(* IEC 61131-3 sources: ZPLC/tools/hil/il_tests, 12 files *)

(* ---- arithmetic.il ---- *)
PROGRAM Arithmetic
VAR
  a AT %QW0 : INT;
  b AT %QW1 : INT;
  res_add AT %QW2 : INT;
  res_sub AT %QW3 : INT;
  res_mul AT %QW4 : INT;
  res_div AT %QW5 : INT;
  res_mod AT %QW6 : INT;
END_VAR

(* Explicit init for test stability *)
LD 10
ST a
LD 5
ST b

LD a
ADD b
ST res_add
LD a
SUB b
ST res_sub
LD a
MUL b
ST res_mul
LD a
DIV b
ST res_div
LD a
MOD b
ST res_mod
END_PROGRAM

(* ---- basic_il.il ---- *)
PROGRAM ILTest
VAR
    a AT %QW0 : INT := 10;
    b AT %QW1 : INT := 20;
    res AT %QW2 : INT;
    flag AT %QX6.0 : BOOL;
END_VAR

LD a
ADD b
ST res

LD res
GT 25
ST flag

END_PROGRAM

(* ---- blinky.il ---- *)
PROGRAM BlinkIL
VAR
  Blink : TON;
  Led AT %QX0.0 : BOOL;
END_VAR

(* The timer runs while the LED is off. When it is done the LED is on for one scan, which restarts the timer. *)
  LDN Led
  ST Blink.IN
  CAL Blink(PT := T#200ms)
  LD Blink.Q
  ST Led
END_PROGRAM

(* ---- comparison.il ---- *)
PROGRAM Comparison
VAR
  val AT %QW0 : INT;
  is_gt AT %QX2.0 : BOOL;
  is_lt AT %QX3.0 : BOOL;
  is_eq AT %QX4.0 : BOOL;
  is_ne AT %QX5.0 : BOOL;
END_VAR

(* Explicit init *)
LD 50
ST val

LD val
GT 40
ST is_gt

LD val
LT 60
ST is_lt

LD val
EQ 50
ST is_eq

LD val
NE 99
ST is_ne
END_PROGRAM

(* ---- debug_bool.il ---- *)
PROGRAM DebugBool
VAR
  res_true AT %QX0.0 : BOOL;
  res_false AT %QX0.1 : BOOL;
END_VAR

LD TRUE
ST res_true

LD FALSE
ST res_false
END_PROGRAM

(* ---- debug_bool.st ---- *)
PROGRAM DebugBool
VAR
  res_true AT %QX0.0 : BOOL;
  res_false AT %QX0.1 : BOOL;
END_VAR

VAR
    IL_CR : DINT;
    IL_CR_BOOL : BOOL;
    IL_CR_REAL : REAL;
END_VAR

(* Test Direct True Load *)
IL_CR_BOOL := TRUE;
res_true := IL_CR_BOOL;

(* Test Direct False Load *)
IL_CR_BOOL := FALSE;
res_false := IL_CR_BOOL;

END_PROGRAM

(* ---- debug_gt.il ---- *)
PROGRAM DebugGT
VAR
  res_gt AT %QX0.0 : BOOL;
END_VAR

LD 50
GT 40
ST res_gt
END_PROGRAM

(* ---- debug_manual.st ---- *)
PROGRAM ILTest
VAR
    a AT %QW0 : INT := 10;
    b AT %QW1 : INT := 20;
    res AT %QW2 : INT;
    flag AT %QX6.0 : BOOL;
END_VAR
VAR
    IL_CR : DINT;
    IL_CR_BOOL : BOOL;
    IL_CR_REAL : REAL;
END_VAR

    IL_CR_BOOL := a <> 0;
    IL_CR := BOOL_TO_INT(IL_CR_BOOL);
END_PROGRAM

(* ---- debug_var.il ---- *)
PROGRAM DebugVar
VAR
  val AT %QW0 : INT;
  res_gt AT %QX2.0 : BOOL;
END_VAR

LD 50
ST val

LD val
GT 40
ST res_gt
END_PROGRAM

(* ---- jumps.il ---- *)
PROGRAM Jumps
VAR
  (* Results - all should stay at their initial values *)
  skip1_result AT %QW0 : INT := 0;
  skip2_result AT %QW1 : INT := 0;
  exec1_result AT %QW2 : INT := 0;
  exec2_result AT %QW3 : INT := 0;
  jump_cond AT %QX8.0 : BOOL := TRUE;
END_VAR

(* Test 1: JMPC - Conditional Jump when TRUE *)
(* When jump_cond is TRUE, skip the next code *)
LD jump_cond
JMPC AfterSkip1

(* This should be SKIPPED when jump_cond=TRUE *)
LD 999
ST skip1_result

AfterSkip1:
(* This always executes - set exec1_result to 42 *)
LD 42
ST exec1_result

(* Test 2: JMP - Unconditional Jump *)
JMP AfterSkip2

(* This should ALWAYS be skipped *)
LD 888
ST skip2_result

AfterSkip2:
(* This always executes - set exec2_result to 77 *)
LD 77
ST exec2_result

END_PROGRAM

(* ---- logic.il ---- *)
PROGRAM Logic
VAR
  t AT %QX0.0 : BOOL := TRUE;
  f AT %QX1.0 : BOOL := FALSE;
  res_and AT %QX2.0 : BOOL;
  res_or AT %QX3.0 : BOOL;
  res_xor AT %QX4.0 : BOOL;
  res_not AT %QX5.0 : BOOL;
END_VAR

(* Explicit Init *)
LD TRUE
ST t
LD FALSE
ST f

LD t
AND f
ST res_and

LD t
OR f
ST res_or

LD t
XOR f
ST res_xor

LD t
NOT
ST res_not
END_PROGRAM

(* ---- minimal.il ---- *)
PROGRAM Minimal
VAR
  res AT %QW0 : INT;
END_VAR
LD 123
ST res
END_PROGRAM
